(* IEC 61131-3 sources: plc-vscode/tests/st/all/trust-platform/crates/trust-runtime/tests/fixtures/oscat/core/src/24_device_driver, 1 file *)

(* ---- tests.st ---- *)
TEST_PROGRAM oscat_device_driver_switching_helpers_behave
VAR
    Driver : DRIVER_1;
    Driver4 : DRIVER_4;
    Driver4C : DRIVER_4C;
    Flow : FLOW_CONTROL;
END_VAR

Driver(SET_REQ := FALSE, IN := FALSE, RST := TRUE, Timeout := T#0s, Toggle_Mode := FALSE);
ASSERT_FALSE(IN := Driver.Q);
Driver(SET_REQ := FALSE, IN := TRUE, RST := FALSE, Timeout := T#0s, Toggle_Mode := FALSE);
ASSERT_TRUE(IN := Driver.Q);
Driver(SET_REQ := FALSE, IN := FALSE, RST := TRUE, Timeout := T#0s, Toggle_Mode := FALSE);
ASSERT_FALSE(IN := Driver.Q);

Driver4(SET_REQ := FALSE, IN0 := TRUE, IN1 := FALSE, IN2 := FALSE, IN3 := FALSE, RST := FALSE, Toggle_Mode := FALSE, Timeout := T#0s);
ASSERT_TRUE(IN := Driver4.Q0);
ASSERT_FALSE(IN := Driver4.Q1);

Driver4C(IN := TRUE, RST := FALSE, Timeout := T#0s);
ASSERT_EQUAL(EXPECTED := INT#1, ACTUAL := Driver4C.SN);
ASSERT_TRUE(IN := Driver4C.Q0);
ASSERT_FALSE(IN := Driver4C.Q1);

Flow(IN := TRUE, REQ := FALSE, ENQ := TRUE, RST := FALSE, T_AUTO := T#0s, T_DELAY := T#0s);
ASSERT_TRUE(IN := Flow.Q);
ASSERT_EQUAL(EXPECTED := BYTE#101, ACTUAL := Flow.STATUS);
END_TEST_PROGRAM

TEST_PROGRAM oscat_device_driver_interlocks_and_manuals_behave
VAR
    Lock2 : INTERLOCK;
    Lock4 : INTERLOCK_4;
    Manual1 : MANUAL_1;
    Manual2 : MANUAL_2;
    Manual4 : MANUAL_4;
END_VAR

Lock2(I1 := TRUE, I2 := FALSE, TL := T#0s);
ASSERT_TRUE(IN := Lock2.Q1);
ASSERT_FALSE(IN := Lock2.Q2);

Lock4(I0 := FALSE, I1 := TRUE, I2 := TRUE, I3 := FALSE, E := TRUE, MODE := INT#1);
ASSERT_EQUAL(EXPECTED := BYTE#4, ACTUAL := Lock4.OUT);
ASSERT_TRUE(IN := Lock4.TP);

ASSERT_TRUE(IN := MANUAL(IN := TRUE, FORCE_ON := FALSE, FORCE_OFF := FALSE));
ASSERT_FALSE(IN := MANUAL(IN := TRUE, FORCE_ON := FALSE, FORCE_OFF := TRUE));

Manual1(IN := FALSE, MAN := TRUE, M_I := TRUE, SET_REQ := FALSE, RST := FALSE);
ASSERT_TRUE(IN := Manual1.Q);
ASSERT_EQUAL(EXPECTED := BYTE#103, ACTUAL := Manual1.STATUS);

Manual2(IN := FALSE, ENA := TRUE, FORCE_ON := TRUE, FORCE_OFF := FALSE, MAN := FALSE);
ASSERT_TRUE(IN := Manual2.Q);
ASSERT_EQUAL(EXPECTED := BYTE#101, ACTUAL := Manual2.STATUS);

Manual4(I0 := FALSE, I1 := FALSE, I2 := FALSE, I3 := FALSE, MAN := TRUE, STP := FALSE, M0 := TRUE, M1 := FALSE, M2 := TRUE, M3 := FALSE);
ASSERT_TRUE(IN := Manual4.Q0);
ASSERT_FALSE(IN := Manual4.Q1);
ASSERT_TRUE(IN := Manual4.Q2);
ASSERT_FALSE(IN := Manual4.Q3);
END_TEST_PROGRAM

TEST_PROGRAM oscat_device_driver_parameter_helpers_behave
VAR
    Pset : PARSET;
    Pset2 : PARSET2;
END_VAR

Pset(A0 := FALSE, A1 := FALSE, X01 := REAL#1.0, X02 := REAL#2.0, X03 := REAL#3.0, X04 := REAL#4.0, X11 := REAL#10.0, X12 := REAL#20.0, X13 := REAL#30.0, X14 := REAL#40.0, X21 := REAL#100.0, X22 := REAL#200.0, X23 := REAL#300.0, X24 := REAL#400.0, X31 := REAL#1000.0, X32 := REAL#2000.0, X33 := REAL#3000.0, X34 := REAL#4000.0, TC := T#0s);
ASSERT_NEAR(EXPECTED := REAL#1.0, ACTUAL := Pset.P1, DELTA := REAL#0.001);
Pset(A0 := TRUE, A1 := FALSE, X01 := REAL#1.0, X02 := REAL#2.0, X03 := REAL#3.0, X04 := REAL#4.0, X11 := REAL#10.0, X12 := REAL#20.0, X13 := REAL#30.0, X14 := REAL#40.0, X21 := REAL#100.0, X22 := REAL#200.0, X23 := REAL#300.0, X24 := REAL#400.0, X31 := REAL#1000.0, X32 := REAL#2000.0, X33 := REAL#3000.0, X34 := REAL#4000.0, TC := T#0s);
ASSERT_NEAR(EXPECTED := REAL#10.0, ACTUAL := Pset.P1, DELTA := REAL#0.001);
Pset(A0 := FALSE, A1 := TRUE, X01 := REAL#1.0, X02 := REAL#2.0, X03 := REAL#3.0, X04 := REAL#4.0, X11 := REAL#10.0, X12 := REAL#20.0, X13 := REAL#30.0, X14 := REAL#40.0, X21 := REAL#100.0, X22 := REAL#200.0, X23 := REAL#300.0, X24 := REAL#400.0, X31 := REAL#1000.0, X32 := REAL#2000.0, X33 := REAL#3000.0, X34 := REAL#4000.0, TC := T#0s);
ASSERT_NEAR(EXPECTED := REAL#100.0, ACTUAL := Pset.P1, DELTA := REAL#0.001);

Pset2(X := REAL#0.5, X01 := REAL#1.0, X02 := REAL#2.0, X03 := REAL#3.0, X04 := REAL#4.0, X11 := REAL#10.0, X12 := REAL#20.0, X13 := REAL#30.0, X14 := REAL#40.0, X21 := REAL#100.0, X22 := REAL#200.0, X23 := REAL#300.0, X24 := REAL#400.0, X31 := REAL#1000.0, X32 := REAL#2000.0, X33 := REAL#3000.0, X34 := REAL#4000.0, L1 := REAL#1.0, L2 := REAL#2.0, L3 := REAL#3.0, TC := T#0s);
ASSERT_NEAR(EXPECTED := REAL#1.0, ACTUAL := Pset2.P1, DELTA := REAL#0.001);
Pset2(X := REAL#1.5, X01 := REAL#1.0, X02 := REAL#2.0, X03 := REAL#3.0, X04 := REAL#4.0, X11 := REAL#10.0, X12 := REAL#20.0, X13 := REAL#30.0, X14 := REAL#40.0, X21 := REAL#100.0, X22 := REAL#200.0, X23 := REAL#300.0, X24 := REAL#400.0, X31 := REAL#1000.0, X32 := REAL#2000.0, X33 := REAL#3000.0, X34 := REAL#4000.0, L1 := REAL#1.0, L2 := REAL#2.0, L3 := REAL#3.0, TC := T#0s);
ASSERT_NEAR(EXPECTED := REAL#10.0, ACTUAL := Pset2.P1, DELTA := REAL#0.001);
Pset2(X := REAL#2.5, X01 := REAL#1.0, X02 := REAL#2.0, X03 := REAL#3.0, X04 := REAL#4.0, X11 := REAL#10.0, X12 := REAL#20.0, X13 := REAL#30.0, X14 := REAL#40.0, X21 := REAL#100.0, X22 := REAL#200.0, X23 := REAL#300.0, X24 := REAL#400.0, X31 := REAL#1000.0, X32 := REAL#2000.0, X33 := REAL#3000.0, X34 := REAL#4000.0, L1 := REAL#1.0, L2 := REAL#2.0, L3 := REAL#3.0, TC := T#0s);
ASSERT_NEAR(EXPECTED := REAL#100.0, ACTUAL := Pset2.P1, DELTA := REAL#0.001);
Pset2(X := REAL#3.5, X01 := REAL#1.0, X02 := REAL#2.0, X03 := REAL#3.0, X04 := REAL#4.0, X11 := REAL#10.0, X12 := REAL#20.0, X13 := REAL#30.0, X14 := REAL#40.0, X21 := REAL#100.0, X22 := REAL#200.0, X23 := REAL#300.0, X24 := REAL#400.0, X31 := REAL#1000.0, X32 := REAL#2000.0, X33 := REAL#3000.0, X34 := REAL#4000.0, L1 := REAL#1.0, L2 := REAL#2.0, L3 := REAL#3.0, TC := T#0s);
ASSERT_NEAR(EXPECTED := REAL#1000.0, ACTUAL := Pset2.P1, DELTA := REAL#0.001);
END_TEST_PROGRAM

TEST_PROGRAM oscat_device_driver_tuning_helpers_behave
VAR
    Ramp : SRAMP;
    FineTune : TUNE;
    FastTune : TUNE2;
    Encoder : INC_DEC;
END_VAR

Ramp(X := REAL#10.0, A_UP := REAL#1.0, A_DN := REAL#-1.0, VU_MAX := REAL#5.0, VD_MAX := REAL#-5.0, LIMIT_HIGH := REAL#100.0, LIMIT_LOW := REAL#0.0, RST := TRUE);
ASSERT_NEAR(EXPECTED := REAL#0.0, ACTUAL := Ramp.Y, DELTA := REAL#0.001);
ASSERT_NEAR(EXPECTED := REAL#0.0, ACTUAL := Ramp.V, DELTA := REAL#0.001);

FineTune(SET_REQ := TRUE, SU := FALSE, SD := FALSE, RST := FALSE, LIMIT_L := REAL#0.0, LIMIT_H := REAL#100.0, RST_val := REAL#5.0, SET_val := REAL#25.0);
ASSERT_NEAR(EXPECTED := REAL#25.0, ACTUAL := FineTune.Y, DELTA := REAL#0.001);
FineTune(SET_REQ := FALSE, SU := FALSE, SD := FALSE, RST := TRUE, LIMIT_L := REAL#0.0, LIMIT_H := REAL#100.0, RST_val := REAL#5.0, SET_val := REAL#25.0);
ASSERT_NEAR(EXPECTED := REAL#5.0, ACTUAL := FineTune.Y, DELTA := REAL#0.001);

FastTune(SET_REQ := TRUE, SU := FALSE, SD := FALSE, FU := FALSE, FD := FALSE, RST := FALSE, LIMIT_L := REAL#0.0, LIMIT_H := REAL#100.0, RST_val := REAL#7.0, SET_val := REAL#30.0);
ASSERT_NEAR(EXPECTED := REAL#30.0, ACTUAL := FastTune.Y, DELTA := REAL#0.001);
FastTune(SET_REQ := FALSE, SU := FALSE, SD := FALSE, FU := FALSE, FD := FALSE, RST := TRUE, LIMIT_L := REAL#0.0, LIMIT_H := REAL#100.0, RST_val := REAL#7.0, SET_val := REAL#30.0);
ASSERT_NEAR(EXPECTED := REAL#7.0, ACTUAL := FastTune.Y, DELTA := REAL#0.001);

Encoder(CHa := FALSE, CHb := FALSE, RST := TRUE);
ASSERT_EQUAL(EXPECTED := INT#0, ACTUAL := Encoder.cnt);
Encoder(CHa := TRUE, CHb := FALSE, RST := FALSE);
ASSERT_TRUE(IN := Encoder.dir);
ASSERT_EQUAL(EXPECTED := INT#1, ACTUAL := Encoder.cnt);
END_TEST_PROGRAM
